(* IEC 61131-3 sources: COMPLCconexMQTT/plcnext_st, 6 files *)

(* ---- PRG_Alarms.st ---- *)
(* ============================================================================
   PROGRAMA: PRG_Alarms
   ENTORNO : Phoenix Contact PLCnext Engineer 2026.6 (AXC F 2152)
   OBJETIVO: Gestión centralizada de alarmas (sensor, comunicación, actuador,
             comando inválido) y restablecimiento controlado por flanco.
   ============================================================================ *)
PROGRAM PRG_Alarms
VAR_EXTERNAL
    SYS_Alarm           : BOOL;   (* Alarma activa general *)
    CMD_Reset_Alarm     : BOOL;   (* Comando remoto de reset *)
    DIAG_Last_Error     : STRING;
END_VAR

VAR_INPUT
    xSensor_Fault       : BOOL;
    xComm_Lost_Alarm    : BOOL;
    xActuator_Fault     : BOOL;
    xInvalid_Cmd_Alarm  : BOOL;
    xInput_Fault        : BOOL;
    xLocal_Reset        : BOOL := FALSE;
END_VAR

VAR_OUTPUT
    xAlarm_Latched      : BOOL;
    xAny_Fault_Active   : BOOL;
END_VAR

VAR
    fbRTRIG_Remote_Rst  : R_TRIG;
    fbRTRIG_Local_Rst   : R_TRIG;
    xReset_Pulse        : BOOL;
END_VAR

(* 1. Evaluar fallas activas *)
xAny_Fault_Active := xSensor_Fault OR xComm_Lost_Alarm OR xActuator_Fault OR xInvalid_Cmd_Alarm OR xInput_Fault;

(* 2. Enclavamiento de alarma *)
IF xAny_Fault_Active THEN
    xAlarm_Latched := TRUE;
END_IF;

(* 3. Detección de flanco de restablecimiento *)
fbRTRIG_Remote_Rst(CLK := CMD_Reset_Alarm);
fbRTRIG_Local_Rst(CLK := xLocal_Reset);
xReset_Pulse := fbRTRIG_Remote_Rst.Q OR fbRTRIG_Local_Rst.Q;

(* Limpiar comando remoto tipo pulso después de procesarlo *)
IF CMD_Reset_Alarm THEN
    CMD_Reset_Alarm := FALSE;
END_IF;

(* 4. Restablecimiento controlado: solo si ya no hay falla física/comunicación *)
IF xReset_Pulse THEN
    IF NOT xAny_Fault_Active THEN
        xAlarm_Latched  := FALSE;
        DIAG_Last_Error := 'OK_ALARM_RESET';
    ELSE
        DIAG_Last_Error := 'WARN_RESET_REJECTED_FAULT_ACTIVE';
    END_IF;
END_IF;

SYS_Alarm := xAlarm_Latched;

END_PROGRAM

(* ---- PRG_Analog.st ---- *)
(* ============================================================================
   PROGRAMA: PRG_Analog
   ENTORNO : Phoenix Contact PLCnext Engineer 2026.6 (AXC F 2152)
   OBJETIVO: Lectura de sensor analógico 0-10 V, conversión a voltaje y %,
             filtrado digital exponencial y validación de rango.
   NOTA    : Ajustar rRaw_Min / rRaw_Max según la hoja de datos del módulo
             Axioline F AI real una vez identificado (ej. 0..30000 en AXL F).
   ============================================================================ *)
PROGRAM PRG_Analog
VAR_EXTERNAL
    AI_Sensor_Raw       : DINT;   (* Valor crudo del módulo analógico *)
    AI_Sensor_Voltage   : REAL;   (* Voltaje calculado [0.0 .. 10.0 V] *)
    AI_Sensor_Percent   : REAL;   (* Porcentaje escalado [0.0 .. 100.0 %] *)
    SYS_Sensor_Valid    : BOOL;   (* TRUE si la lectura está dentro de rango válido *)
    DIAG_Last_Error     : STRING;
END_VAR

VAR_INPUT
    diRaw_Min           : DINT := 0;      (* Ajustar según módulo AXL F real *)
    diRaw_Max           : DINT := 30000;  (* Ajustar según módulo AXL F real *)
    rFilter_Alpha       : REAL := 0.2;    (* Factor de filtro EMA (0.05 .. 1.0) *)
    rVoltage_Min_Valid  : REAL := -0.2;   (* Tolerancia inferior de cero *)
    rVoltage_Max_Valid  : REAL := 10.5;   (* Tolerancia superior de sobre-rango *)
END_VAR

VAR_OUTPUT
    xSensor_Fault       : BOOL;
END_VAR

VAR
    rSpan               : REAL;
    rVoltage_Raw        : REAL;
    rVoltage_Filtered   : REAL := 0.0;
    xFirst_Scan         : BOOL := TRUE;
    rAlpha_Clamped      : REAL;
END_VAR

(* 1. Validar parámetros de escalamiento *)
rSpan := DINT_TO_REAL(diRaw_Max - diRaw_Min);
IF rSpan <= 0.0 THEN
    SYS_Sensor_Valid := FALSE;
    xSensor_Fault    := TRUE;
    DIAG_Last_Error  := 'FAULT_ANALOG_CONFIG_SPAN';
    RETURN;
END_IF;

(* 2. Conversión lineal crudo -> Voltaje (0-10 V) *)
rVoltage_Raw := (DINT_TO_REAL(AI_Sensor_Raw - diRaw_Min) / rSpan) * 10.0;

(* 3. Validación de rango y detección de valores anormales / rotura / corto *)
IF (rVoltage_Raw < rVoltage_Min_Valid) OR (rVoltage_Raw > rVoltage_Max_Valid) THEN
    SYS_Sensor_Valid := FALSE;
    xSensor_Fault    := TRUE;
    DIAG_Last_Error  := 'FAULT_SENSOR_OUT_OF_RANGE';
ELSE
    SYS_Sensor_Valid := TRUE;
    xSensor_Fault    := FALSE;
END_IF;

(* 4. Limitar voltaje físico para cálculo limpio [0.0 .. 10.0 V] *)
IF rVoltage_Raw < 0.0 THEN
    rVoltage_Raw := 0.0;
ELSIF rVoltage_Raw > 10.0 THEN
    rVoltage_Raw := 10.0;
END_IF;

(* 5. Filtro digital exponencial configurable (EMA) *)
rAlpha_Clamped := rFilter_Alpha;
IF rAlpha_Clamped < 0.01 THEN rAlpha_Clamped := 0.01; END_IF;
IF rAlpha_Clamped > 1.0  THEN rAlpha_Clamped := 1.0;  END_IF;

IF xFirst_Scan THEN
    rVoltage_Filtered := rVoltage_Raw;
    xFirst_Scan       := FALSE;
ELSE
    rVoltage_Filtered := (rAlpha_Clamped * rVoltage_Raw) + ((1.0 - rAlpha_Clamped) * rVoltage_Filtered);
END_IF;

(* 6. Publicación de salidas *)
AI_Sensor_Voltage := rVoltage_Filtered;
AI_Sensor_Percent := (AI_Sensor_Voltage / 10.0) * 100.0;

END_PROGRAM

(* ---- PRG_Communication.st ---- *)
(* ============================================================================
   PROGRAMA: PRG_Communication
   ENTORNO : Phoenix Contact PLCnext Engineer 2026.6 (AXC F 2152)
   OBJETIVO: Heartbeat del PLC, monitoreo de Heartbeat del Gateway (Node-RED)
             con watchdog configurable y recuperación segura sin arranques.
   ============================================================================ *)
PROGRAM PRG_Communication
VAR_EXTERNAL
    SYS_PLC_Heartbeat       : UDINT; (* Contador incremental del PLC (cada 1 s) *)
    SYS_Gateway_Heartbeat   : UDINT; (* Contador escrito por Node-RED vía OPC UA *)
    SYS_Communication_OK    : BOOL;  (* TRUE = Gateway activo dentro del watchdog *)
    DIAG_OPC_UA_Status      : BOOL;  (* Estado lógico de enlace OPC UA *)
    DIAG_Last_Error         : STRING;
END_VAR

VAR_INPUT
    tHeartbeat_Period       : TIME := T#1s;
    tWatchdog_Timeout       : TIME := T#5s;
END_VAR

VAR_OUTPUT
    xComm_Lost_Alarm        : BOOL;
    xComm_Restored_Pulse    : BOOL;
END_VAR

VAR
    fbTON_PLC_HB            : TON;
    fbTON_Watchdog          : TON;
    udiLast_Gateway_HB      : UDINT := 0;
    xFirst_Scan             : BOOL := TRUE;
    xPrev_Comm_OK           : BOOL := FALSE;
    fbRTRIG_Comm_OK         : R_TRIG;
END_VAR

(* 1. Generación de Heartbeat del PLC (1 Hz) *)
fbTON_PLC_HB(IN := NOT fbTON_PLC_HB.Q, PT := tHeartbeat_Period);
IF fbTON_PLC_HB.Q THEN
    SYS_PLC_Heartbeat := SYS_PLC_Heartbeat + 1;
END_IF;

(* 2. Watchdog sobre el Heartbeat del Gateway *)
IF xFirst_Scan THEN
    udiLast_Gateway_HB := SYS_Gateway_Heartbeat;
    xFirst_Scan        := FALSE;
END_IF;

IF SYS_Gateway_Heartbeat <> udiLast_Gateway_HB THEN
    (* Hubo actividad nueva del Gateway: reiniciar watchdog *)
    udiLast_Gateway_HB := SYS_Gateway_Heartbeat;
    fbTON_Watchdog(IN := FALSE, PT := tWatchdog_Timeout);
    SYS_Communication_OK := TRUE;
    DIAG_OPC_UA_Status   := TRUE;
    xComm_Lost_Alarm     := FALSE;
ELSE
    fbTON_Watchdog(IN := TRUE, PT := tWatchdog_Timeout);
    IF fbTON_Watchdog.Q THEN
        SYS_Communication_OK := FALSE;
        DIAG_OPC_UA_Status   := FALSE;
        xComm_Lost_Alarm     := TRUE;
        DIAG_Last_Error      := 'ALARM_COMM_WATCHDOG_TIMEOUT';
    END_IF;
END_IF;

(* 3. Pulso de recuperación (solo informativo; NO genera orden de marcha) *)
fbRTRIG_Comm_OK(CLK := SYS_Communication_OK);
xComm_Restored_Pulse := fbRTRIG_Comm_OK.Q;
xPrev_Comm_OK        := SYS_Communication_OK;

END_PROGRAM

(* ---- PRG_Inputs.st ---- *)
(* ============================================================================
   PROGRAMA: PRG_Inputs
   ENTORNO : Phoenix Contact PLCnext Engineer 2026.6 (AXC F 2152)
   OBJETIVO: Lectura de entradas digitales (Start / Stop) con antirrebote,
             detección de flancos y diagnóstico básico de entradas.
   NOTA    : Mapear DI_Start_Raw y DI_Stop_Raw en Port List cuando se
             identifique el módulo Axioline F real (NO inventar direcciones).
   ============================================================================ *)
PROGRAM PRG_Inputs
VAR_EXTERNAL
    DI_Start            : BOOL;   (* Pulsador de arranque filtrado (NA) *)
    DI_Stop             : BOOL;   (* Pulsador de parada filtrado *)
    DIAG_Last_Error     : STRING; (* Último mensaje de diagnóstico *)
END_VAR

VAR_INPUT
    xRaw_Start          : BOOL;   (* Enlazar a canal DI físico del módulo AXL F *)
    xRaw_Stop           : BOOL;   (* Enlazar a canal DI físico del módulo AXL F *)
    xStop_Is_NC         : BOOL := FALSE; (* TRUE si el pulsador físico Stop es NC *)
    tDebounce_Time      : TIME := T#50ms;
END_VAR

VAR_OUTPUT
    xStart_Pulse        : BOOL;   (* Flanco ascendente de arranque válido *)
    xStop_Active        : BOOL;   (* TRUE = condición de parada activa *)
    xInput_Fault        : BOOL;   (* Falla por pulsación simultánea prolongada *)
END_VAR

VAR
    fbTON_Start         : TON;
    fbTON_Stop          : TON;
    fbTON_Both_Pressed  : TON;
    fbRTRIG_Start       : R_TRIG;
    xStop_Normalized    : BOOL;
END_VAR

(* 1. Normalización de lógica NC/NA para el pulsador de parada *)
IF xStop_Is_NC THEN
    xStop_Normalized := NOT xRaw_Stop;
ELSE
    xStop_Normalized := xRaw_Stop;
END_IF;

(* 2. Filtrado antirrebote *)
fbTON_Start(IN := xRaw_Start, PT := tDebounce_Time);
fbTON_Stop(IN := xStop_Normalized, PT := tDebounce_Time);

DI_Start := fbTON_Start.Q;
DI_Stop  := fbTON_Stop.Q;

(* 3. Detección de flanco para arranque *)
fbRTRIG_Start(CLK := DI_Start);
xStart_Pulse := fbRTRIG_Start.Q;
xStop_Active := DI_Stop;

(* 4. Diagnóstico: Start y Stop activos simultáneamente > 2 s *)
fbTON_Both_Pressed(IN := (DI_Start AND DI_Stop), PT := T#2s);
xInput_Fault := fbTON_Both_Pressed.Q;

IF xInput_Fault THEN
    DIAG_Last_Error := 'FAULT_INPUTS_SIMULTANEOUS_START_STOP';
END_IF;

END_PROGRAM

(* ---- PRG_Main.st ---- *)
(* ============================================================================
   PROGRAMA: PRG_Main
   ENTORNO : Phoenix Contact PLCnext Engineer 2026.6 (AXC F 2152)
   OBJETIVO: Programa principal coordinador y declaración de variables globales
             compartidas con OPC UA.
   ============================================================================ *)
PROGRAM PRG_Main
VAR
    (* Entradas físicas / simbólicas *)
    DI_Start                : BOOL := FALSE;
    DI_Stop                 : BOOL := FALSE;
    AI_Sensor_Raw           : DINT := 0;
    AI_Sensor_Voltage       : REAL := 0.0;
    AI_Sensor_Percent       : REAL := 0.0;

    (* Salidas físicas / simbólicas *)
    DO_Motor                : BOOL := FALSE;
    DO_LED                  : BOOL := FALSE;

    (* Comandos remotos OPC UA (Lectura/Escritura) *)
    CMD_Motor_Start         : BOOL := FALSE;
    CMD_Motor_Stop          : BOOL := FALSE;
    CMD_LED                 : BOOL := FALSE;
    CMD_Reset_Alarm         : BOOL := FALSE;

    (* Estado del sistema *)
    SYS_PLC_Heartbeat       : UDINT := 0;
    SYS_Gateway_Heartbeat   : UDINT := 0;
    SYS_Communication_OK    : BOOL := FALSE;
    SYS_Motor_Status        : BOOL := FALSE;
    SYS_Alarm               : BOOL := FALSE;
    SYS_Sensor_Valid        : BOOL := FALSE;
    SYS_System_Ready        : BOOL := FALSE;

    (* Diagnóstico *)
    DIAG_OPC_UA_Status      : BOOL := FALSE;
    DIAG_MQTT_Status        : BOOL := FALSE;
    DIAG_Last_Command_ID    : STRING := '';
    DIAG_Last_Error         : STRING := '';

    (* Instancias de subprogramas *)
    instInputs              : PRG_Inputs;
    instAnalog              : PRG_Analog;
    instComm                : PRG_Communication;
    instAlarms              : PRG_Alarms;
    instMotor               : PRG_Motor;
END_VAR

(* 1. Lectura y filtrado de entradas digitales *)
instInputs();

(* 2. Lectura y escalamiento analógico 0-10 V *)
instAnalog();

(* 3. Watchdog y Heartbeats *)
instComm();

(* 4. Estado listo del sistema *)
SYS_System_Ready := (NOT SYS_Alarm) AND SYS_Sensor_Valid;

(* 5. Control del motor *)
instMotor(
    xLocal_Start_Pulse := instInputs.xStart_Pulse,
    xLocal_Stop_Active := instInputs.xStop_Active
);

(* 6. Gestión centralizada de alarmas *)
instAlarms(
    xSensor_Fault      := instAnalog.xSensor_Fault,
    xComm_Lost_Alarm   := instComm.xComm_Lost_Alarm,
    xActuator_Fault    := instMotor.xActuator_Fault,
    xInvalid_Cmd_Alarm := instMotor.xInvalid_Cmd_Alarm,
    xInput_Fault       := instInputs.xInput_Fault
);

END_PROGRAM

(* ---- PRG_Motor.st ---- *)
(* ============================================================================
   PROGRAMA: PRG_Motor
   ENTORNO : Phoenix Contact PLCnext Engineer 2026.6 (AXC F 2152)
   OBJETIVO: Control local y remoto del motor con prioridad de parada física,
             validación de permisos, enclavamiento y control de LED indicador.
   ============================================================================ *)
PROGRAM PRG_Motor
VAR_EXTERNAL
    DO_Motor                : BOOL;   (* Salida física hacia contactor/motor *)
    DO_LED                  : BOOL;   (* Salida física LED indicador *)
    CMD_Motor_Start         : BOOL;   (* Comando remoto de arranque *)
    CMD_Motor_Stop          : BOOL;   (* Comando remoto de parada *)
    CMD_LED                 : BOOL;   (* Comando remoto de LED *)
    SYS_Communication_OK    : BOOL;
    SYS_Motor_Status        : BOOL;
    SYS_Alarm               : BOOL;
    SYS_Sensor_Valid        : BOOL;
    SYS_System_Ready        : BOOL;
    DIAG_Last_Command_ID    : STRING;
    DIAG_Last_Error         : STRING;
END_VAR

VAR_INPUT
    xLocal_Start_Pulse      : BOOL;   (* Flanco de pulsador físico Start *)
    xLocal_Stop_Active      : BOOL;   (* Pulsador físico Stop (PRIORIDAD 1) *)
    xMotor_Feedback         : BOOL := TRUE; (* Opcional: realimentación contactor *)
    xUse_Feedback           : BOOL := FALSE;
    tFeedback_Timeout       : TIME := T#2s;
END_VAR

VAR_OUTPUT
    xActuator_Fault         : BOOL;
    xInvalid_Cmd_Alarm      : BOOL;
END_VAR

VAR
    fbRTRIG_Remote_Start    : R_TRIG;
    fbRTRIG_Remote_Stop     : R_TRIG;
    fbTON_Feedback          : TON;
    xMotor_Latch            : BOOL := FALSE;
    xRemote_Start_Allowed   : BOOL;
END_VAR

(* 1. Detección de flancos de comandos remotos *)
fbRTRIG_Remote_Start(CLK := CMD_Motor_Start);
fbRTRIG_Remote_Stop(CLK := CMD_Motor_Stop);

(* 2. Condición de permiso para comandos remotos *)
xRemote_Start_Allowed := SYS_Communication_OK AND SYS_System_Ready AND (NOT SYS_Alarm) AND SYS_Sensor_Valid;

(* 3. PRIORIDAD 1: Parada física o parada remota o alarma crítica *)
IF xLocal_Stop_Active OR fbRTRIG_Remote_Stop.Q OR SYS_Alarm THEN
    xMotor_Latch := FALSE;
END_IF;

(* 4. Arranque local (siempre permitido si no hay Stop físico ni alarma) *)
IF xLocal_Start_Pulse AND (NOT xLocal_Stop_Active) AND (NOT SYS_Alarm) THEN
    xMotor_Latch := TRUE;
END_IF;

(* 5. Arranque remoto (sujeto a permisos y sin Stop físico) *)
IF fbRTRIG_Remote_Start.Q THEN
    IF xRemote_Start_Allowed AND (NOT xLocal_Stop_Active) THEN
        xMotor_Latch := TRUE;
    ELSE
        xInvalid_Cmd_Alarm := TRUE;
        DIAG_Last_Error    := 'CMD_REMOTE_START_REJECTED_INTERLOCK';
    END_IF;
END_IF;

(* 6. Limpiar comandos remotos tras ser evaluados (evita re-arranques al reconectar) *)
IF CMD_Motor_Start THEN
    CMD_Motor_Start := FALSE;
END_IF;
IF CMD_Motor_Stop THEN
    CMD_Motor_Stop := FALSE;
END_IF;

(* 7. Asignación de salidas físicas *)
DO_Motor         := xMotor_Latch;
SYS_Motor_Status := DO_Motor;

(* LED: encendido si motor activo o si comando remoto de LED está activo y hay comunicación *)
DO_LED := DO_Motor OR (CMD_LED AND SYS_Communication_OK);

(* 8. Diagnóstico opcional de realimentación de contactor *)
IF xUse_Feedback THEN
    fbTON_Feedback(IN := (DO_Motor <> xMotor_Feedback), PT := tFeedback_Timeout);
    xActuator_Fault := fbTON_Feedback.Q;
    IF xActuator_Fault THEN
        xMotor_Latch    := FALSE;
        DO_Motor        := FALSE;
        DIAG_Last_Error := 'FAULT_ACTUATOR_FEEDBACK_MISMATCH';
    END_IF;
ELSE
    xActuator_Fault := FALSE;
END_IF;

END_PROGRAM
